(* IEC 61131-3 sources: plc-process-lib/tests/POUs/Suites/FB_Integration_Test, 9 files *)

(* ---- AiPidVfdTracksBumplessNoWindup.method.decl.st ---- *)
// Контур уровня КНС по примеру 17.3 контракта: LT (AI 4–20 мА, 0..10 м) -> LIC (ПИД Direct, Kp 2, Ti 20 с,
// xUseOutAct) -> ведущий насос (ПЧ, rSpeedMin 30 %); xTrack := NOT SpeedAutoActive, rTrack = rOutAct = SpeedRef с
// прошлого цикла. (1) Насос стоит в Auto — ПИД следит, выход = заданию ПЧ (0 %), Available = FALSE. (2) Пуск:
// Starting — ПИД ещё следит (30 % — предустановка ПЧ); Running — слежение снято, выход ПИД без рывка (30 %).
// (3) Уровень 4,8 м ниже задания 5 м 10 мин: ПИД просит меньше минимума, задание ПЧ держится на 30 %, выход ПИД по
// обратному расчёту от rOutAct не уходит в 0: 30 + P = 30 - 2·2 = 26 %. (4) Уровень 5,2 м — задание ПЧ сразу 34 %
// (30 + P), без задержки на «раскрутку» интегратора.
METHOD PRIVATE AiPidVfdTracksBumplessNoWindup
VAR
    fbTime   : FB_FakeTime;          // подменное время, старт 1 ч
    fbAi     : FB_AnalogInput;       // LT: уровень 4–20 мА, 0..10 м
    stAiCmd  : ST_AnalogInputCmd;    // его команды
    stAiCfg  : ST_AnalogInputCfg;    // его Cfg
    fbPid    : FB_PID;               // LIC: регулятор уровня
    stPidCmd : ST_PidCmd;            // его команды
    stPidRet : ST_DeviceRetain;      // его режим
    stPidCfg : ST_PidCfg;            // его Cfg
    fbVfd    : FB_MotorVfd;          // ведущий насос с ПЧ
    stVfdCmd : ST_MotorCmd;          // его команды
    stVfdRet : ST_DeviceRetain;      // его режим и счётчики
    stVfdCfg : ST_MotorCfg;          // его Cfg
END_VAR

(* ---- AllTypesAlarmCountThroughIDevice.method.decl.st ---- *)
// Все семь типов доступны через I_Device (интерфейс станции и SCADA-адаптера): число слотов тревог
// AlarmCount (I_AlarmSource) после первого вызова равно <DEV>_ALARM_COUNT из GVL_Const, слот 0
// доступен через GetAlarm, режим — из перечисления. У FB_Motor и FB_MotorVfd слотов одинаково (8).
METHOD PRIVATE AllTypesAlarmCountThroughIDevice
VAR
    fbTime   : FB_FakeTime;          // подменное время, старт 1 ч
    fbAi     : FB_AnalogInput;       // аналоговый вход
    stAiCmd  : ST_AnalogInputCmd;    // его команды
    stAiCfg  : ST_AnalogInputCfg;    // его Cfg (умолчания)
    fbDi     : FB_DigitalInput;      // дискретный вход
    stDiCmd  : ST_DigitalInputCmd;   // его команды
    stDiCfg  : ST_DigitalInputCfg;   // его Cfg (умолчания)
    fbMot    : FB_Motor;             // двигатель прямого пуска
    stMotCmd : ST_MotorCmd;          // его команды
    stMotRet : ST_DeviceRetain;      // его retain
    stMotCfg : ST_MotorCfg;          // его Cfg (умолчания)
    fbVfd    : FB_MotorVfd;          // двигатель с ПЧ
    stVfdCmd : ST_MotorCmd;          // его команды
    stVfdRet : ST_DeviceRetain;      // его retain
    stVfdCfg : ST_MotorCfg;          // его Cfg (умолчания, с полем stVfd)
    fbVlv    : FB_Valve;             // запорная арматура
    stVlvCmd : ST_ValveCmd;          // её команды
    stVlvRet : ST_DeviceRetain;      // её retain
    stVlvCfg : ST_ValveCfg;          // её Cfg (умолчания)
    fbCv     : FB_ControlValve;      // регулирующий клапан
    stCvCmd  : ST_ControlValveCmd;   // его команды
    stCvRet  : ST_DeviceRetain;      // его retain
    stCvCfg  : ST_ControlValveCfg;   // его Cfg (умолчания)
    fbPid    : FB_PID;               // ПИД-регулятор
    stPidCmd : ST_PidCmd;            // его команды
    stPidRet : ST_DeviceRetain;      // его retain
    stPidCfg : ST_PidCfg;            // его Cfg (умолчания)
    aitfDev  : ARRAY[1..7] OF I_Device;   // устройства через интерфейс
    auiSlots : ARRAY[1..7] OF UINT;       // ожидаемое число слотов
    uiDev    : UINT;                      // номер устройства
    itfAlm   : I_Alarm;                   // слот 0 устройства
    xCountOk : BOOL := TRUE;              // у всех AlarmCount совпал
    xSlotOk  : BOOL := TRUE;              // у всех слот 0 доступен
    xModeOk  : BOOL := TRUE;              // у всех режим из перечисления
END_VAR

(* ---- AllTypesAlarmCountThroughIDevice.method.impl.st ---- *)
coUnit.TEST('Device_AllTypes_AlarmCountThroughIDevice');

fbAi(itfTime := fbTime, stCmd := stAiCmd, stCfg := stAiCfg);
fbDi(itfTime := fbTime, stCmd := stDiCmd, stCfg := stDiCfg);
fbMot(itfTime := fbTime, stCmd := stMotCmd, stRetain := stMotRet, stCfg := stMotCfg);
fbVfd(itfTime := fbTime, stCmd := stVfdCmd, stRetain := stVfdRet, stCfg := stVfdCfg);
fbVlv(itfTime := fbTime, stCmd := stVlvCmd, stRetain := stVlvRet, stCfg := stVlvCfg);
fbCv(itfTime := fbTime, stCmd := stCvCmd, stRetain := stCvRet, stCfg := stCvCfg);
fbPid(itfTime := fbTime, stCmd := stPidCmd, stRetain := stPidRet, stCfg := stPidCfg);
aitfDev[1] := fbAi;
aitfDev[2] := fbDi;
aitfDev[3] := fbMot;
aitfDev[4] := fbVfd;
aitfDev[5] := fbVlv;
aitfDev[6] := fbCv;
aitfDev[7] := fbPid;
auiSlots[1] := GVL_Const.AI_ALARM_COUNT;
auiSlots[2] := GVL_Const.DI_ALARM_COUNT;
auiSlots[3] := GVL_Const.MOT_ALARM_COUNT;
auiSlots[4] := GVL_Const.MOT_ALARM_COUNT;
auiSlots[5] := GVL_Const.VLV_ALARM_COUNT;
auiSlots[6] := GVL_Const.CV_ALARM_COUNT;
auiSlots[7] := GVL_Const.PID_ALARM_COUNT;
FOR uiDev := 1 TO 7 DO
    xCountOk := xCountOk AND (aitfDev[uiDev].AlarmCount = auiSlots[uiDev]);
    itfAlm := aitfDev[uiDev].GetAlarm(uiIndex := 0);
    xSlotOk := xSlotOk AND (itfAlm <> 0);
    xModeOk := xModeOk AND (aitfDev[uiDev].Mode = E_DeviceMode.Auto OR aitfDev[uiDev].Mode = E_DeviceMode.Manual
                            OR aitfDev[uiDev].Mode = E_DeviceMode.Local
                            OR aitfDev[uiDev].Mode = E_DeviceMode.OutOfService);
END_FOR
AssertTrue(Condition := xCountOk, Message := 'AlarmCount = <DEV>_ALARM_COUNT for every type');
AssertTrue(Condition := xSlotOk, Message := 'slot 0 reachable through GetAlarm');
AssertTrue(Condition := xModeOk, Message := 'mode from the enumeration');
AssertEquals_UINT(Expected := GVL_Const.MOT_ALARM_COUNT, Actual := fbVfd.AlarmCount,
                  Message := 'MotorVfd: eight slots like Motor');

coUnit.TEST_FINISHED();

(* ---- DefaultCfgPassesCheck.method.decl.st ---- *)
// Инвариант генератора (контракт 2.3, раздел 20): умолчания Cfg всех семи типов устройств проходят
// CheckConfig — после первого вызова wCfgErr = 0 и нет бита DEV_STS_CFG_ERROR (корректная Cfg принята
// как LKG). Каждый тип — настоящий ФБ, а не тестовое устройство (F-26).
METHOD PRIVATE DefaultCfgPassesCheck
VAR
    fbTime   : FB_FakeTime;          // подменное время, старт 1 ч
    fbAi     : FB_AnalogInput;       // аналоговый вход
    stAiCmd  : ST_AnalogInputCmd;    // его команды
    stAiCfg  : ST_AnalogInputCfg;    // его Cfg (умолчания)
    fbDi     : FB_DigitalInput;      // дискретный вход
    stDiCmd  : ST_DigitalInputCmd;   // его команды
    stDiCfg  : ST_DigitalInputCfg;   // его Cfg (умолчания)
    fbMot    : FB_Motor;             // двигатель прямого пуска
    stMotCmd : ST_MotorCmd;          // его команды
    stMotRet : ST_DeviceRetain;      // его retain
    stMotCfg : ST_MotorCfg;          // его Cfg (умолчания)
    fbVfd    : FB_MotorVfd;          // двигатель с ПЧ
    stVfdCmd : ST_MotorCmd;          // его команды
    stVfdRet : ST_DeviceRetain;      // его retain
    stVfdCfg : ST_MotorCfg;          // его Cfg (умолчания, с полем stVfd)
    fbVlv    : FB_Valve;             // запорная арматура
    stVlvCmd : ST_ValveCmd;          // её команды
    stVlvRet : ST_DeviceRetain;      // её retain
    stVlvCfg : ST_ValveCfg;          // её Cfg (умолчания)
    fbCv     : FB_ControlValve;      // регулирующий клапан
    stCvCmd  : ST_ControlValveCmd;   // его команды
    stCvRet  : ST_DeviceRetain;      // его retain
    stCvCfg  : ST_ControlValveCfg;   // его Cfg (умолчания)
    fbPid    : FB_PID;               // ПИД-регулятор
    stPidCmd : ST_PidCmd;            // его команды
    stPidRet : ST_DeviceRetain;      // его retain
    stPidCfg : ST_PidCfg;            // его Cfg (умолчания)
END_VAR

(* ---- DevTypeReportedInStsCommon.method.decl.st ---- *)
// Каждый тип пишет свой E_DeviceType в stSts.stCommon.eDevType с первого вызова (SCADA выбирает
// фейсплейт, генератор карты Modbus сверяет тип блока); до первого вызова — None. FB_MotorVfd
// сообщает MotorVfd, а не Motor: FB_Motor тип наследника не затирает и во втором вызове.
METHOD PRIVATE DevTypeReportedInStsCommon
VAR
    fbTime   : FB_FakeTime;          // подменное время, старт 1 ч
    fbAi     : FB_AnalogInput;       // аналоговый вход
    stAiCmd  : ST_AnalogInputCmd;    // его команды
    stAiCfg  : ST_AnalogInputCfg;    // его Cfg (умолчания)
    fbDi     : FB_DigitalInput;      // дискретный вход
    stDiCmd  : ST_DigitalInputCmd;   // его команды
    stDiCfg  : ST_DigitalInputCfg;   // его Cfg (умолчания)
    fbMot    : FB_Motor;             // двигатель прямого пуска
    stMotCmd : ST_MotorCmd;          // его команды
    stMotRet : ST_DeviceRetain;      // его retain
    stMotCfg : ST_MotorCfg;          // его Cfg (умолчания)
    fbVfd    : FB_MotorVfd;          // двигатель с ПЧ
    stVfdCmd : ST_MotorCmd;          // его команды
    stVfdRet : ST_DeviceRetain;      // его retain
    stVfdCfg : ST_MotorCfg;          // его Cfg (умолчания, с полем stVfd)
    fbVlv    : FB_Valve;             // запорная арматура
    stVlvCmd : ST_ValveCmd;          // её команды
    stVlvRet : ST_DeviceRetain;      // её retain
    stVlvCfg : ST_ValveCfg;          // её Cfg (умолчания)
    fbCv     : FB_ControlValve;      // регулирующий клапан
    stCvCmd  : ST_ControlValveCmd;   // его команды
    stCvRet  : ST_DeviceRetain;      // его retain
    stCvCfg  : ST_ControlValveCfg;   // его Cfg (умолчания)
    fbPid    : FB_PID;               // ПИД-регулятор
    stPidCmd : ST_PidCmd;            // его команды
    stPidRet : ST_DeviceRetain;      // его retain
    stPidCfg : ST_PidCfg;            // его Cfg (умолчания)
END_VAR

(* ---- GuardBandCurrentPidHoldsOutput.method.decl.st ---- *)
// Датчик уровня выдаёт ток отказа NAMUR, а канал AI читает 3,61 мА (защитная полоса NE 43, AI-13). ПИД (Reverse,
// Auto, задание 5 м, выход 40 %) работает tFailDelay = 2 с по значению насыщения, затем AI снимает xValid — ПИД
// фиксирует отказ PV и удерживает выход (Hold), а не уводит его к 100 % за минуту.
METHOD PRIVATE GuardBandCurrentPidHoldsOutput
VAR
    fbTime   : FB_FakeTime;          // подменное время, старт 1 ч
    fbAi     : FB_AnalogInput;       // LT: уровень 4–20 мА, 0..10 м
    stAiCmd  : ST_AnalogInputCmd;    // его команды
    stAiCfg  : ST_AnalogInputCfg;    // его Cfg
    fbPid    : FB_PID;               // LIC: регулятор уровня
    stPidCmd : ST_PidCmd;            // его команды
    stPidRet : ST_DeviceRetain;      // его режим
    stPidCfg : ST_PidCfg;            // его Cfg
    iStep    : INT;                  // шаг цикла
    rOut5s   : REAL;                 // выход ПИД через 5 с
END_VAR

(* ---- GuardBandCurrentPidHoldsOutput.method.impl.st ---- *)
coUnit.TEST('LevelLoop_GuardBandCurrent_PidHoldsOutput');

stAiCfg.rRangeHi_eu := 10.0;
stPidCfg.rPvMax_eu := 10.0;
stPidCfg.rSpMax_eu := 10.0;
stPidRet.eRemoteMode := E_DeviceMode.Auto;
stPidCmd.rSp_eu := 5.0;
stPidCmd.rManualOut_pct := 40.0;
FOR iStep := 1 TO 600 DO
    fbTime.Advance(tStep := T#100MS);
    fbAi(itfTime := fbTime, rIn := 3.61, stCmd := stAiCmd, stCfg := stAiCfg);
    fbPid(itfTime := fbTime, rPv_eu := fbAi.rValue_eu, xPvValid := fbAi.xValid, stCmd := stPidCmd,
          stRetain := stPidRet, stCfg := stPidCfg);
    IF iStep = 50 THEN
        rOut5s := fbPid.rOut_pct;
    END_IF
END_FOR
AssertFalse(Condition := fbAi.xValid, Message := 'guard band confirmed: PV invalid');
AssertEquals_WORD(Expected := GVL_Const.PID_FLT_PV_INVALID, Actual := fbPid.stSts.stCommon.wFault,
                  Message := 'PID reports the PV fault');
AssertTrue(Condition := fbPid.rOut_pct < 50.0, Message := 'output held, not driven to 100 pct');
AssertEquals_REAL(Expected := rOut5s, Actual := fbPid.rOut_pct, Delta := 1.0E-4,
                  Message := 'output frozen after the fault');

coUnit.TEST_FINISHED();

(* ---- LevelLoopStep.method.decl.st ---- *)
// Помощник: uiN циклов контура уровня по примеру 17.3 контракта, перед каждым — шаг подменного времени tDt
// (T#0S — тот же момент): ведущий насос (прошлый вызов) -> AI -> ПИД (xTrack := NOT SpeedAutoActive,
// rTrack = rOutAct = SpeedRef) -> задание ПЧ -> ПЧ -> модель ПЧ (работает по команде, скорость = заданию).
// Ассертов внутри нет
METHOD PRIVATE LevelLoopStep
VAR_IN_OUT
    fbT      : FB_FakeTime;          // подменное время
    fbAi     : FB_AnalogInput;       // датчик уровня
    stAiCmd  : ST_AnalogInputCmd;    // его команды
    fbPid    : FB_PID;               // регулятор уровня
    stPidCmd : ST_PidCmd;            // его команды
    stPidRet : ST_DeviceRetain;      // его режим
    fbVfd    : FB_MotorVfd;          // ведущий насос
    stVfdCmd : ST_MotorCmd;          // его команды
    stVfdRet : ST_DeviceRetain;      // его режим и счётчики
END_VAR
VAR_IN_OUT CONSTANT
    stAiCfg  : ST_AnalogInputCfg;    // Cfg датчика
    stPidCfg : ST_PidCfg;            // Cfg регулятора
    stVfdCfg : ST_MotorCfg;          // Cfg насоса
END_VAR
VAR_INPUT
    rLevel_mA : REAL;                // ток датчика уровня, мА
    uiN       : UINT;                // число циклов
    tDt       : TIME;                // шаг времени перед каждым циклом
END_VAR
VAR
    uiLoop    : UINT;                // номер цикла
    xLeadAuto : BOOL;                // ведущий насос в Auto и работает (прошлый цикл)
    rLeadRef  : REAL;                // задание ведущего насоса (прошлый цикл), %
END_VAR

(* ---- LevelLoopStep.method.impl.st ---- *)
FOR uiLoop := 1 TO uiN DO
    fbT.Advance(tStep := tDt);
    xLeadAuto := fbVfd.SpeedAutoActive;
    rLeadRef := fbVfd.SpeedRef;
    fbAi(itfTime := fbT, rIn := rLevel_mA, stCmd := stAiCmd, stCfg := stAiCfg);
    fbPid(itfTime := fbT, rPv_eu := fbAi.rValue_eu, xPvValid := fbAi.xValid, xTrack := NOT xLeadAuto,
          rTrack_pct := rLeadRef, rOutAct_pct := rLeadRef, stCmd := stPidCmd, stRetain := stPidRet, stCfg := stPidCfg);
    fbVfd.rSpeedSpAuto_pct := fbPid.rOut_pct;
    fbVfd(itfTime := fbT, stCmd := stVfdCmd, stRetain := stVfdRet, stCfg := stVfdCfg);
    fbVfd.xVfdRunning := fbVfd.xQRun;
    fbVfd.rSpeedAct_pct := SEL(fbVfd.xQRun, 0.0, fbVfd.rSpeedRef_pct);
END_FOR
